(* IEC 61131-3 sources: ZPLC/packages/zplc-ide/plant-scenes/buffer-release, 2 files *)

(* ---- reference.st ---- *)
PROGRAM BufferRelease
VAR_INPUT
    Start      AT %I0.0 : BOOL;
    ReleaseCmd AT %I0.1 : BOOL;
    EyeFull    AT %I0.2 : BOOL;
    EyeBlade   AT %I0.3 : BOOL;
    EyeRelease AT %I0.4 : BOOL;
END_VAR
VAR_OUTPUT
    RunBuffer  AT %Q0.0 : BOOL;
    RunRelease AT %Q0.1 : BOOL;
    Emit       AT %Q0.2 : BOOL;
    Hold       AT %Q0.3 : BOOL;
    Done       AT %Q0.4 : BOOL;
    Fault      AT %Q0.5 : BOOL;
END_VAR
VAR
    Active    : BOOL;
    Releasing : BOOL;
    Pace      : TON;
    Loaded    : CTU;
    Cmd       : R_TRIG;
    Passed    : F_TRIG;
    Entered   : R_TRIG;
    Sent      : CTU;
    Extra     : BOOL;
END_VAR

IF Start THEN
    Active := TRUE;
END_IF;

(* load: one box every two seconds until five are on the belt *)
Pace(IN := Active AND NOT Pace.Q AND NOT Loaded.Q, PT := T#2s);
Emit := Pace.Q;
Loaded(CU := Pace.Q, R := FALSE, PV := 5);

(* release: one box per command, the blade stays down until that box has passed EyeRelease *)
Cmd(CLK := ReleaseCmd);
Entered(CLK := EyeRelease);
Passed(CLK := EyeRelease);
IF Cmd.Q AND Loaded.Q AND EyeBlade AND NOT Releasing THEN
    Releasing := TRUE;
END_IF;
(* a box reaching EyeRelease with no command pending means a second box got through *)
IF Entered.Q AND NOT Releasing THEN
    Extra := TRUE;
END_IF;
IF Releasing AND Passed.Q THEN
    Releasing := FALSE;
END_IF;
Sent(CU := Passed.Q, R := FALSE, PV := 5);

Hold := Active AND NOT Releasing;
(* the buffer belt waits while a box is released, so the next box cannot follow it *)
RunBuffer := Active AND NOT Releasing;
RunRelease := Active;
Done := Sent.Q;
Fault := Extra;

END_PROGRAM

(* ---- starter.st ---- *)
PROGRAM BufferRelease
VAR_INPUT
    Start      AT %I0.0 : BOOL;  (* StartButton.pressed: start loading the buffer *)
    ReleaseCmd AT %I0.1 : BOOL;  (* ReleaseButton.pressed: one press releases one box *)
    EyeFull    AT %I0.2 : BOOL;  (* EyeFull.detect: sees the fifth box in the queue *)
    EyeBlade   AT %I0.3 : BOOL;  (* EyeBlade.detect: sees the box waiting at the blade *)
    EyeRelease AT %I0.4 : BOOL;  (* EyeRelease.detect: sees each box that leaves the blade *)
END_VAR
VAR_OUTPUT
    RunBuffer  AT %Q0.0 : BOOL;  (* Buffer1.run: run the buffer belt *)
    RunRelease AT %Q0.1 : BOOL;  (* Release1.run: run the release belt *)
    Emit       AT %Q0.2 : BOOL;  (* Emitter1.emit: put one box on the buffer belt *)
    Hold       AT %Q0.3 : BOOL;  (* Blade1.extend: the blade holds the queue while true *)
    Done       AT %Q0.4 : BOOL;  (* DoneLight.lit: lit when five boxes have been released *)
    Fault      AT %Q0.5 : BOOL;  (* FaultLight.lit: lit if a release lets a second box through *)
END_VAR

(* Goal: a press of the start button loads five boxes, one every two seconds,
   and the blade holds them in a queue. Each press of the release button
   lowers the blade just long enough for one box to pass EyeRelease, then
   raises it again. Light Done after the fifth box, and Fault if a release
   ever lets two boxes through. *)

END_PROGRAM
